Fanuc KAREL source: kd00027.KL

-- PROVISIONAL review KL for V1013-1; original PC SHA256 8d4737db122d9bfedfd6a6ce348acb79c9d2452400cfb141d00f033f8a364e4f
-- Incomplete behavior may be omitted. Consult companion uncertainty JSON. Do not deploy.
PROGRAM KD00027
%NOLOCKGROUP
VAR
  I : INTEGER
  J : INTEGER
  B : BOOLEAN
  R : REAL
  S : STRING[80]
BEGIN
  -- UNRESOLVED_PC offsets 5-21; opcodes 9D,81,18,9D,12,22,9D,13,04
  -- UNRESOLVED_PC offsets 26-30; opcodes 7F
END KD00027
